// TIA Portal V21 export
// export: Created 2026-10-14T03:11:21.1521181Z, ExportSetting WithDefaults, DisplayName Totally Integrated Automation Portal, DisplayVersion V21, DisplayName STEP 7 Professional, DisplayVersion V21, DisplayName STEP 7 Safety, DisplayVersion V21, DisplayName Tech WebApplication, DisplayVersion V21, DisplayName WinCC Basic/Comfort/Advanced, DisplayVersion V21, DisplayName WinCC Unified, DisplayVersion V21
TagTable "AccError"
  LLCCA_ErrAcc_DB_LLCCA_PID_oErrAcc : LReal  (HMI_Connection_1, 100 ms)
  LLCCA_ErrAcc_DB_PID_C_oErrAcc : LReal  (HMI_Connection_1, 100 ms)
